Fanuc KAREL source: kt00259.KL

-- PROVISIONAL review KL for V770-1; original PC SHA256 fbfbb40c0176aa47ba80632696dd948e8b3b1fa4aff784a181ba7f25d68c2dee
-- Incomplete behavior may be omitted. Consult companion uncertainty JSON. Do not deploy.
PROGRAM KT00259
%NOLOCKGROUP
VAR
  I1 : INTEGER
  OUT : BOOLEAN
-- UNRESOLVED_DECL Y2 type=002018
BEGIN
  -- UNRESOLVED_PC offsets 5-16; opcodes 2E,23
  -- UNRESOLVED_PC offsets 21-35; opcodes 2E,22,9D,33,B2
  -- UNRESOLVED_PC offsets 40-62; opcodes 21,22,9D,33,B1,57,23
  -- UNRESOLVED_PC offsets 67-71; opcodes 7F
END KT00259
